(* IEC 61131-3 sources: dvigatel_dorosh/codesys, 10 files *)

(* ---- 00_DUT_MotorTypes.st ---- *)
TYPE E_MotorState :
(
    MOTOR_DISABLED,
    MOTOR_IDLE,
    MOTOR_RAMP,
    MOTOR_WAIT_STOP,
    MOTOR_RUN,
    MOTOR_FAULT
);
END_TYPE

TYPE ST_MotorCommand :
STRUCT
    SpeedRPM : REAL;
    RampSec : REAL;
    Direction : INT; // +1 / -1
    Sequence : WORD;
END_STRUCT
END_TYPE

(* ---- 01_GVL_PC.st ---- *)
VAR_GLOBAL
    // Explicitly map these words into Modbus TCP holding registers in Device Tree.
    // 0..5: PC request. 100..116: PLC telemetry.
    Holding : ARRAY[0..127] OF WORD;

    // Must be commissioned ON SITE; no automatic activation from Ethernet.
    CommissionEnable : BOOL := FALSE;
    ConfigValid : BOOL := FALSE;
    PGFeedbackProven : BOOL := FALSE;
    HardwareSafetyOK : BOOL := FALSE;

    // Assign IO in device mappings, not hard-coded addresses.
    Pt100TemperatureC : REAL;
    Pt100InputValid : BOOL;
END_VAR

(* ---- 07_GVL_DriveIO.st ---- *)
VAR_GLOBAL
    // Link via CODESYS Modbus Serial Device I/O Mapping.
    // NEVER assume default values mean communication is healthy.
    SpeedRaw : WORD;
    StatusRaw : WORD;
    FrequencyRaw : WORD;
    CurrentRaw : WORD;
    FaultCodeRaw : WORD;
    SpeedResponsePulse : BOOL;
    StatusResponsePulse : BOOL;
    DriveReadFresh : BOOL;
    DriveFault : BOOL;

    // Final outputs are NOT directly mapped to a write device in this version.
    // Implement an acknowledged, single-in-flight Modbus RTU scheduler.
    PendingFrequencyWord : WORD;
    PendingControlWord : WORD;
END_VAR

(* ---- 02_FB_Pt100Protection.st ---- *)
FUNCTION_BLOCK FB_Pt100Protection
VAR_INPUT
    TemperatureC : REAL;
    ChannelHealthy : BOOL;
    WarningC : REAL;
    TripC : REAL;
    ResetBelowC : REAL;
    Ack : BOOL;
    LimitsConfigured : BOOL;
END_VAR
VAR_OUTPUT
    Warning : BOOL;
    TripLatched : BOOL;
    Valid : BOOL;
    Permit : BOOL;
END_VAR

Valid := ChannelHealthy AND LimitsConfigured
         AND (ResetBelowC < WarningC)
         AND (WarningC < TripC);
Warning := Valid AND (TemperatureC >= WarningC);

IF (NOT Valid) OR (TemperatureC >= TripC) THEN
    TripLatched := TRUE;
END_IF;

// Acknowledgement alone cannot clear fault if input is missing.
IF Ack AND Valid AND (TemperatureC <= ResetBelowC) THEN
    TripLatched := FALSE;
END_IF;
Permit := Valid AND NOT TripLatched;
END_FUNCTION_BLOCK

(* ---- 03_FB_Heartbeat.st ---- *)
FUNCTION_BLOCK FB_Heartbeat
VAR_INPUT
    Counter : WORD;
    Enable : BOOL;
    CycleSec : REAL;
    TimeoutSec : REAL;
END_VAR
VAR_OUTPUT
    Active : BOOL;
END_VAR
VAR
    Previous : WORD;
    AgeSec : REAL := 10000.0;
    Initialized : BOOL;
END_VAR

IF NOT Enable THEN
    Active := FALSE;
    Initialized := FALSE;
    AgeSec := TimeoutSec;
ELSE
    IF NOT Initialized THEN
        Previous := Counter;
        Initialized := TRUE;
        AgeSec := TimeoutSec;
    ELSIF Counter <> Previous THEN
        Previous := Counter;
        AgeSec := 0.0;
    ELSE
        AgeSec := MIN(10000.0, AgeSec + CycleSec);
    END_IF;
    Active := AgeSec < TimeoutSec;
END_IF;
END_FUNCTION_BLOCK

(* ---- 04_FB_ConfirmedStop.st ---- *)
FUNCTION_BLOCK FB_ConfirmedStop
VAR_INPUT
    EncoderFeedbackProven : BOOL;
    SpeedFresh : BOOL;
    StatusFresh : BOOL;
    DriveReportsStopped : BOOL;
    MeasuredRPM : REAL;
    CycleSec : REAL;
    ThresholdRPM : REAL;
    StableSec : REAL;
END_VAR
VAR_OUTPUT
    Confirmed : BOOL;
END_VAR
VAR
    StableForSec : REAL;
END_VAR

IF EncoderFeedbackProven AND SpeedFresh AND StatusFresh
   AND DriveReportsStopped
   AND (ABS(MeasuredRPM) <= ThresholdRPM)
   AND (StableSec > 0.0) THEN
    StableForSec := MIN(StableSec, StableForSec + CycleSec);
ELSE
    StableForSec := 0.0;
END_IF;
Confirmed := StableForSec >= StableSec AND StableSec > 0.0;
END_FUNCTION_BLOCK

(* ---- 05_FB_MotorMotion.st ---- *)
FUNCTION_BLOCK FB_MotorMotion
VAR_INPUT
    Enable : BOOL;
    InterlocksOK : BOOL;
    CommandPulse : BOOL;
    Command : ST_MotorCommand;
    FaultAck : BOOL;
    StopConfirmed : BOOL;
    CycleSec : REAL;
    MaxRPM : REAL;
    StopTimeoutSec : REAL;
END_VAR
VAR_OUTPUT
    State : E_MotorState := MOTOR_DISABLED;
    ProfileRPM : REAL;             // signed reference
    RunRequest : BOOL;
    ReverseRequest : BOOL;
    StopRequest : BOOL := TRUE;
    FaultLatched : BOOL;
    AcceptedSequence : WORD;
END_VAR
VAR
    Goal : REAL;
    StageStart : REAL;
    StageEnd : REAL;
    StageSec : REAL;
    StageAge : REAL;
    StopAge : REAL;
    PendingReverse : BOOL;
    HeldDirection : INT := 1;
    NewGoal : BOOL;
    ValidCmd : BOOL;
END_VAR

// Device safety must NOT depend on a functioning serial link.
// This output requests a controlled stop; hardware safety is separate.
IF NOT Enable THEN
    State := MOTOR_DISABLED;
    ProfileRPM := 0.0;
    Goal := 0.0;
    PendingReverse := FALSE;
ELSIF NOT InterlocksOK THEN
    FaultLatched := TRUE;
    State := MOTOR_FAULT;
END_IF;

IF State = MOTOR_FAULT THEN
    // Explicit acknowledgement while truly stopped. Does not re-launch.
    IF FaultAck AND InterlocksOK AND StopConfirmed
       AND (Command.SpeedRPM = 0.0) AND NOT CommandPulse THEN
        FaultLatched := FALSE;
        State := MOTOR_IDLE;
        ProfileRPM := 0.0;
        Goal := 0.0;
    END_IF;
ELSIF State = MOTOR_DISABLED THEN
    // Moving from disabled to idle does not accept any pre-existing command.
    IF Enable AND InterlocksOK AND StopConfirmed THEN
        State := MOTOR_IDLE;
    END_IF;
ELSIF Enable AND InterlocksOK THEN
    ValidCmd := (Command.Direction = 1 OR Command.Direction = -1)
            AND (Command.SpeedRPM >= 0.0)
            AND (Command.SpeedRPM <= MaxRPM)
            AND (Command.RampSec >= 0.1)
            AND (Command.RampSec <= 600.0)
            AND (MaxRPM > 0.0);

    NewGoal := CommandPulse AND ValidCmd;
    IF NewGoal THEN
        AcceptedSequence := Command.Sequence;
        Goal := Command.SpeedRPM * INT_TO_REAL(Command.Direction);
        StageSec := Command.RampSec;

        IF State = MOTOR_WAIT_STOP THEN
            // Never cancel physical-stop gate on a new command.
            PendingReverse := (ABS(Goal) > 0.001);
        ELSE
            StageStart := ProfileRPM;
            StageAge := 0.0;
            IF (ABS(ProfileRPM) > 0.001) AND (ABS(Goal) > 0.001)
               AND ((ProfileRPM > 0.0) <> (Goal > 0.0)) THEN
                StageEnd := 0.0;    // reverse: first stop
                PendingReverse := TRUE;
            ELSIF (ABS(ProfileRPM) < 0.001) AND (NOT StopConfirmed)
                  AND (ABS(Goal) > 0.001) THEN
                State := MOTOR_WAIT_STOP;
                StopAge := 0.0;
                PendingReverse := TRUE;
            ELSE
                StageEnd := Goal;
                PendingReverse := FALSE;
                IF ABS(ProfileRPM) < 0.001 AND ABS(Goal) > 0.001 THEN
                    IF Goal < 0.0 THEN HeldDirection := -1;
                    ELSE HeldDirection := 1; END_IF;
                END_IF;
            END_IF;
            IF State <> MOTOR_WAIT_STOP THEN State := MOTOR_RAMP; END_IF;
        END_IF;
    END_IF;

    CASE State OF
        MOTOR_IDLE:
            ProfileRPM := 0.0;

        MOTOR_RAMP:
            StageAge := MIN(StageSec, StageAge + CycleSec);
            ProfileRPM := StageStart +
                 (StageEnd - StageStart) * (StageAge / StageSec);
            IF StageAge >= StageSec THEN
                ProfileRPM := StageEnd;
                IF ABS(StageEnd) <= 0.001 THEN
                    StopAge := 0.0;
                    State := MOTOR_WAIT_STOP;
                ELSE
                    State := MOTOR_RUN;
                END_IF;
            END_IF;

        MOTOR_WAIT_STOP:
            ProfileRPM := 0.0;
            StopAge := StopAge + CycleSec;
            IF StopConfirmed THEN
                IF ABS(Goal) <= 0.001 THEN
                    PendingReverse := FALSE;
                    State := MOTOR_IDLE;
                ELSE
                    IF Goal < 0.0 THEN HeldDirection := -1;
                    ELSE HeldDirection := 1; END_IF;
                    StageStart := 0.0;
                    StageEnd := Goal;
                    StageAge := 0.0;
                    PendingReverse := FALSE;
                    State := MOTOR_RAMP;
                END_IF;
            ELSIF StopAge >= StopTimeoutSec THEN
                FaultLatched := TRUE;
                State := MOTOR_FAULT;
            END_IF;

        MOTOR_RUN:
            ProfileRPM := Goal;
    END_CASE;
END_IF;

// Enforce a stop request for every blocked or waiting state.
RunRequest := (State = MOTOR_RAMP OR State = MOTOR_RUN)
              AND ABS(ProfileRPM) > 0.001
              AND InterlocksOK AND Enable AND NOT FaultLatched;
ReverseRequest := HeldDirection = -1;
StopRequest := NOT RunRequest;
IF State = MOTOR_FAULT OR State = MOTOR_DISABLED THEN
    ProfileRPM := 0.0;
    RunRequest := FALSE;
    StopRequest := TRUE;
END_IF;
END_FUNCTION_BLOCK

(* ---- 06_FB_DriveCommand.st ---- *)
FUNCTION_BLOCK FB_DriveCommand
VAR_INPUT
    ProfileRPM : REAL;
    RunRequest : BOOL;
    ReverseRequest : BOOL;
    StopRequest : BOOL;
    MotorPolePairs : UINT;
    MaximumHz : REAL;
    ConfigurationValid : BOOL;
END_VAR
VAR_OUTPUT
    FrequencyHz : REAL;
    FrequencyWord : WORD;
    ControlWord : WORD;
    Valid : BOOL;
END_VAR

// Feedforward only: true shaft RPM is read from drive.
// This formula does NOT correct asynchronous slip.
Valid := ConfigurationValid AND (MotorPolePairs > 0)
         AND (MaximumHz > 0.0) AND (MaximumHz <= 300.0);
IF NOT Valid THEN
    FrequencyHz := 0.0;
    FrequencyWord := 0;
    ControlWord := 16#0004; // nominal deceleration-stop candidate; verify at bench
ELSE
    FrequencyHz := LIMIT(0.0,
         ABS(ProfileRPM) * UINT_TO_REAL(MotorPolePairs) / 60.0,
         MaximumHz);
    FrequencyWord := REAL_TO_WORD(FrequencyHz * 100.0);
    IF StopRequest OR NOT RunRequest THEN
        ControlWord := 16#0004;
    ELSIF ReverseRequest THEN
        ControlWord := 16#0003;
    ELSE
        ControlWord := 16#0001;
    END_IF;
END_IF;
END_FUNCTION_BLOCK

(* ---- 09_FB_InnovertRTU.st ---- *)
FUNCTION_BLOCK FB_InnovertRTU
VAR_INPUT
    EnablePort : BOOL;
    ComPortNumber : UDINT; // Must be confirmed on PLC200 hardware; zero disables.
    SlaveId : USINT := 1;
    Baudrate : UDINT := 38400;
    EnableWrites : BOOL;   // FALSE until verified commissioning.
    CommandPermitted : BOOL; // Set only after hardware + PG + Pt100 and TCP watchdog.
    SetFrequency : WORD;    // 0.01 Hz units after checking P00.00.
    SetControl : WORD;      // manual confirms 0x0001 forward, 0x0003 reverse, 0x0004 stop.
    CycleSec : REAL := 0.02;
END_VAR
VAR_OUTPUT
    PortActive : BOOL;
    Busy : BOOL;
    Healthy : BOOL;
    LastError : BOOL;
    ErrorCount : UDINT;
    OkCount : UDINT;
    LastOperation : UINT;
    LastFailedOperation : UINT;
    SpeedRaw : WORD;
    StatusRaw : WORD;
    FrequencyRaw : WORD;
    CurrentRaw : WORD;
    FaultRaw : WORD;
    SpeedFresh : BOOL;
    StatusFresh : BOOL;
    TelemetryFresh : BOOL;
    WriteFrequencyAck : BOOL;
    WriteControlAck : BOOL;
    LastWrittenFrequency : WORD;
    LastWrittenControl : WORD;
END_VAR
VAR
    Com : OCL.COM_Control;
    Request : OCL.MB_SerialRequest;
    State : UINT := 0;
    Step : UINT := 0;
    RequestExecute : BOOL;
    FC : OCL.MB_FC;
    RegisterAddress : UINT;
    Payload : WORD;
    StepAge : REAL;
    SpeedAge : REAL := 10000.0;
    StatusAge : REAL := 10000.0;
    CurrentAge : REAL := 10000.0;
    FaultAge : REAL := 10000.0;
    FrequencyAge : REAL := 10000.0;
    PendingFrequency : WORD;
    PendingControl : WORD;
    HadWriteFrequencyAck : BOOL;
    HadWriteControlAck : BOOL;
    ErrorStreak : UINT;
    WriteEligible : BOOL;
    IsWrite : BOOL;
    ReadyPort : BOOL;
END_VAR

// One FB owns one physical port. Never create a second Modbus COM Port
// on the same RS-485 interface in the CODESYS Device Tree.
SpeedFresh := FALSE;
StatusFresh := FALSE;
TelemetryFresh := FALSE;
WriteFrequencyAck := FALSE;
WriteControlAck := FALSE;
LastError := FALSE;
Busy := (State = 20);
SpeedAge := MIN(10000.0, SpeedAge + CycleSec);
StatusAge := MIN(10000.0, StatusAge + CycleSec);
FrequencyAge := MIN(10000.0, FrequencyAge + CycleSec);
CurrentAge := MIN(10000.0, CurrentAge + CycleSec);
FaultAge := MIN(10000.0, FaultAge + CycleSec);

// Avoid opening unspecified COM ports.
ReadyPort := EnablePort AND (ComPortNumber > 0);
Com(
    xEnable := ReadyPort,
    udiComPort := ComPortNumber,
    udiBaudrate := Baudrate,
    udiByteSize := 8,
    eParity := OCL.COM_PARITY.NONE,
    eStopBit := OCL.COM_STOPBIT.ONE
);
PortActive := Com.xActive AND NOT Com.xError;

// Keep one request FB called EVERY PLC task with a rising-edge Execute.
Request(
    xExecute := RequestExecute,
    tTimeout := T#300MS,
    usiRetry := 0,
    hCom := Com.hCom,
    xIsAsciiMode := FALSE,
    usiSlaveId := SlaveId,
    eFuncCode := FC,
    uiDataAddr := RegisterAddress,
    uiDataCount := 1,
    pData := ADR(Payload),
    szSize := SIZEOF(Payload)
);

IF NOT PortActive THEN
    State := 0;
    Step := 0;
    RequestExecute := FALSE;
    ErrorStreak := 0;
    SpeedAge := 10000.0;
    StatusAge := 10000.0;
    Healthy := FALSE;
ELSE
    CASE State OF
    0: // start from read-only polling every time port activates
        Step := 0;
        State := 10;
    10: // choose next operation; readings are serialized.
        RequestExecute := FALSE;
        Payload := 0;
        FC := OCL.MB_FC.READ_HOLDING_REGISTERS;
        IsWrite := FALSE;
        CASE Step OF
        0: RegisterAddress := 16#8107; // RPM
        1: RegisterAddress := 16#8118; // run status
        2: RegisterAddress := 16#8102; // output frequency
        3: RegisterAddress := 16#810A; // output current
        4: RegisterAddress := 16#812B; // fault code
        5:
            // Writing is NEVER enabled by merely connecting the PLC to a PC.
            WriteEligible := EnableWrites AND CommandPermitted
                           AND Healthy AND (SpeedAge < 0.8)
                           AND (StatusAge < 0.8);
            IF WriteEligible THEN
                PendingFrequency := SetFrequency;
                PendingControl := SetControl;
                Payload := PendingFrequency;
                RegisterAddress := 16#0000;
                FC := OCL.MB_FC.WRITE_SINGLE_REGISTER;
                IsWrite := TRUE;
            ELSE
                Step := 0;
                RegisterAddress := 16#8107;
            END_IF;
        6:
            // Cannot write command without a successfully acked frequency write.
            IF HadWriteFrequencyAck AND EnableWrites AND CommandPermitted THEN
                Payload := PendingControl;
                RegisterAddress := 16#8000;
                FC := OCL.MB_FC.WRITE_SINGLE_REGISTER;
                IsWrite := TRUE;
            ELSE
                Step := 0;
                RegisterAddress := 16#8107;
            END_IF;
        ELSE
            Step := 0;
            RegisterAddress := 16#8107;
        END_CASE;
        LastOperation := Step;
        State := 20;
    20: // Hold execute through busy and until Done or Error
        RequestExecute := TRUE;
        IF Request.xDone THEN
            OkCount := OkCount + 1;
            ErrorStreak := 0;
            IF IsWrite THEN
                IF Step = 5 THEN
                    HadWriteFrequencyAck := TRUE;
                    LastWrittenFrequency := PendingFrequency;
                    WriteFrequencyAck := TRUE;
                ELSIF Step = 6 THEN
                    HadWriteControlAck := TRUE;
                    LastWrittenControl := PendingControl;
                    WriteControlAck := TRUE;
                END_IF;
            ELSE
                CASE Step OF
                0:
                    SpeedRaw := Payload;
                    SpeedAge := 0.0;
                    SpeedFresh := TRUE;
                1:
                    StatusRaw := Payload;
                    StatusAge := 0.0;
                    StatusFresh := TRUE;
                2:
                    FrequencyRaw := Payload;
                    FrequencyAge := 0.0;
                3:
                    CurrentRaw := Payload;
                    CurrentAge := 0.0;
                4:
                    FaultRaw := Payload;
                    FaultAge := 0.0;
                END_CASE;
            END_IF;
            State := 30;
        ELSIF Request.xError THEN
            ErrorCount := ErrorCount + 1;
            LastError := TRUE;
            LastFailedOperation := Step;
            ErrorStreak := ErrorStreak + 1;
            HadWriteFrequencyAck := FALSE;
            HadWriteControlAck := FALSE;
            SpeedAge := 10000.0; // fail closed even if status register still has data
            StatusAge := 10000.0;
            State := 30;
        END_IF;
    30: // create falling edge before next request
        RequestExecute := FALSE;
        State := 40;
    40:
        IF Step >= 6 THEN
            Step := 0;
            HadWriteFrequencyAck := FALSE;
        ELSE
            Step := Step + 1;
        END_IF;
        State := 10;
    END_CASE;
END_IF;

Healthy := PortActive AND (ErrorStreak < 3)
           AND (SpeedAge < 0.8) AND (StatusAge < 0.8);
TelemetryFresh := Healthy AND (FrequencyAge < 2.0)
                  AND (CurrentAge < 2.0) AND (FaultAge < 2.0);
Busy := State = 20;
END_FUNCTION_BLOCK

(* ---- 08_PRG_MotorMain.st ---- *)
PROGRAM PRG_MotorMain
VAR
    // Set PLC_PRG task period to 20 ms and verify actual runtime.
    CycleSec : REAL := 0.02;
    TemperatureWarningC : REAL := 0.0; // configure from motor documentation
    TemperatureTripC : REAL := 0.0;
    TemperatureResetC : REAL := 0.0;
    TemperatureLimitsConfigured : BOOL := FALSE;
    MaximumRPM : REAL := 0.0; // set only after mechanical review
    MaximumHz : REAL := 0.0;
    MotorPolePairs : UINT := 0; // expected 2 for 4 poles, verify
    MaxStopWaitSec : REAL := 30.0;

    // These inputs require proven wiring and runtime diagnostics.
    DriveReportsStopped : BOOL := FALSE;
    DriveStatusDecoded : BOOL := FALSE;
    DriveSpeedScalingProven : BOOL := FALSE;
    DriveSpeedSignedRPM : REAL := 0.0;
    DriveResponseAgeSec : REAL := 10000.0;

    RTU : FB_InnovertRTU;
    RTU_ComPort : UDINT := 0; // Set actual PLC200 COM port from hardware diagnostics
    RTU_WriteEnable : BOOL := FALSE; // Must remain FALSE until commissioning
    Temp : FB_Pt100Protection;
    HB : FB_Heartbeat;
    StopCheck : FB_ConfirmedStop;
    Motion : FB_MotorMotion;
    DriveCmd : FB_DriveCommand;

    Cmd : ST_MotorCommand;
    CmdPulse : BOOL;
    LastRequestID : WORD;
    RequestID : WORD;
    RequestDir : INT;
    ValidRequest : BOOL;
    Interlocks : BOOL;
    RunPermitted : BOOL;
    SpeedFresh : BOOL;
    StatusFresh : BOOL;
    TelemetryState : UINT;
    SignedX10 : DINT;
    SignedX10DW : DWORD;
    Ack : BOOL := FALSE; // safety reset must be engineered separately
END_VAR

// Raw RTU communication: use OwenCommunication library; no Modbus COM Port
// device can occupy the same physical RS-485.
RTU(
    EnablePort:=RTU_ComPort > 0,
    ComPortNumber:=RTU_ComPort,
    SlaveId:=1, Baudrate:=38400,
    EnableWrites:=RTU_WriteEnable,
    CommandPermitted:=RunPermitted,
    SetFrequency:=DriveCmd.FrequencyWord,
    SetControl:=DriveCmd.ControlWord,
    CycleSec:=CycleSec
);
GVL_DriveIO.SpeedRaw := RTU.SpeedRaw;
GVL_DriveIO.StatusRaw := RTU.StatusRaw;
GVL_DriveIO.FrequencyRaw := RTU.FrequencyRaw;
GVL_DriveIO.CurrentRaw := RTU.CurrentRaw;
GVL_DriveIO.FaultCodeRaw := RTU.FaultRaw;
GVL_DriveIO.SpeedResponsePulse := RTU.SpeedFresh;
GVL_DriveIO.StatusResponsePulse := RTU.StatusFresh;
GVL_DriveIO.DriveReadFresh := RTU.Healthy;

// WARNING: The following drive-dependent values must be decoded and proven
// from the real IMD222U21E-ENC diagnostics. Not hardwired to TRUE.
// DriveReportsStopped, DriveStatusDecoded, DriveSpeedScalingProven
// and DriveSpeedSignedRPM are commissioning variables.

// Inputs Holding[0..4] must be protected against concurrent partial writes.
// The application accepts ONLY a changed command ID and validated fields.
// For production replace this elementary transaction handling with a
// verified command buffer / consistency token / single writer.
RequestID := GVL_PC.Holding[4];
RequestDir := 0;
IF GVL_PC.Holding[2] = 1 THEN RequestDir := 1; END_IF;
IF GVL_PC.Holding[2] = 2 THEN RequestDir := -1; END_IF;

Cmd.SpeedRPM := WORD_TO_REAL(GVL_PC.Holding[0]) / 10.0;
Cmd.RampSec := WORD_TO_REAL(GVL_PC.Holding[1]) / 10.0;
Cmd.Direction := RequestDir;
Cmd.Sequence := RequestID;
ValidRequest := RequestDir <> 0
    AND Cmd.SpeedRPM >= 0.0 AND Cmd.SpeedRPM <= MaximumRPM
    AND Cmd.RampSec >= 0.1 AND Cmd.RampSec <= 600.0;

CmdPulse := (RequestID <> LastRequestID) AND ValidRequest;
IF RequestID <> LastRequestID THEN LastRequestID := RequestID; END_IF;

Temp(TemperatureC:=GVL_PC.Pt100TemperatureC,
    ChannelHealthy:=GVL_PC.Pt100InputValid,
    WarningC:=TemperatureWarningC, TripC:=TemperatureTripC,
    ResetBelowC:=TemperatureResetC, Ack:=FALSE,
    LimitsConfigured:=TemperatureLimitsConfigured);
HB(Counter:=GVL_PC.Holding[3], Enable:=GVL_PC.CommissionEnable,
   CycleSec:=CycleSec, TimeoutSec:=2.0);

// Freshness: true pulse must be generated on an actual successful RTU response.
IF GVL_DriveIO.DriveReadFresh THEN
    DriveResponseAgeSec := 0.0;
ELSE
    DriveResponseAgeSec := MIN(10000.0, DriveResponseAgeSec + CycleSec);
END_IF;
SpeedFresh := DriveResponseAgeSec < 0.6 AND DriveSpeedScalingProven
              AND GVL_PC.PGFeedbackProven;
StatusFresh := DriveResponseAgeSec < 0.6 AND DriveStatusDecoded;
StopCheck(EncoderFeedbackProven:=GVL_PC.PGFeedbackProven,
    SpeedFresh:=SpeedFresh, StatusFresh:=StatusFresh,
    DriveReportsStopped:=DriveReportsStopped,
    MeasuredRPM:=DriveSpeedSignedRPM, CycleSec:=CycleSec,
    ThresholdRPM:=5.0, StableSec:=0.4);

RunPermitted := GVL_PC.CommissionEnable AND GVL_PC.ConfigValid
    AND GVL_PC.HardwareSafetyOK AND Temp.Permit AND HB.Active
    AND SpeedFresh AND StatusFresh AND NOT GVL_DriveIO.DriveFault;

Interlocks := RunPermitted;
Motion(Enable:=GVL_PC.CommissionEnable AND GVL_PC.ConfigValid,
    InterlocksOK:=Interlocks,
    CommandPulse:=CmdPulse AND HB.Active, Command:=Cmd,
    FaultAck:=FALSE, StopConfirmed:=StopCheck.Confirmed,
    CycleSec:=CycleSec, MaxRPM:=MaximumRPM,
    StopTimeoutSec:=MaxStopWaitSec);
DriveCmd(ProfileRPM:=Motion.ProfileRPM,
    RunRequest:=Motion.RunRequest,
    ReverseRequest:=Motion.ReverseRequest,
    StopRequest:=Motion.StopRequest,
    MotorPolePairs:=MotorPolePairs, MaximumHz:=MaximumHz,
    ConfigurationValid:=GVL_PC.ConfigValid);

// NOT connected to Modbus write requests by default.
// Once RTU scheduler is implemented, it must send frequency and control
// sequentially, verify each acknowledgement, and latch failures.
GVL_DriveIO.PendingFrequencyWord := DriveCmd.FrequencyWord;
GVL_DriveIO.PendingControlWord := DriveCmd.ControlWord;

CASE Motion.State OF
 MOTOR_DISABLED: TelemetryState := 0;
 MOTOR_IDLE: TelemetryState := 1;
 MOTOR_RAMP: TelemetryState := 2;
 MOTOR_WAIT_STOP: TelemetryState := 3;
 MOTOR_RUN: TelemetryState := 4;
 MOTOR_FAULT: TelemetryState := 90;
END_CASE;

GVL_PC.Holding[100] := Motion.AcceptedSequence;
GVL_PC.Holding[101] := UINT_TO_WORD(TelemetryState);
SignedX10 := REAL_TO_DINT(DriveSpeedSignedRPM * 10.0);
SignedX10DW := DINT_TO_DWORD(SignedX10);
GVL_PC.Holding[102] := DWORD_TO_WORD(SHR(SignedX10DW,16));
GVL_PC.Holding[103] := DWORD_TO_WORD(SignedX10DW AND 16#0000FFFF);
IF GVL_PC.Pt100InputValid THEN
 GVL_PC.Holding[104] := INT_TO_WORD(REAL_TO_INT(GVL_PC.Pt100TemperatureC*10.0));
ELSE
 GVL_PC.Holding[104] := 16#7FFF;
END_IF;
GVL_PC.Holding[105] := GVL_DriveIO.FrequencyRaw;
GVL_PC.Holding[106] := GVL_DriveIO.CurrentRaw;
GVL_PC.Holding[107] := GVL_DriveIO.StatusRaw;
GVL_PC.Holding[108] := GVL_DriveIO.FaultCodeRaw;
GVL_PC.Holding[109] := BOOL_TO_WORD(SpeedFresh AND StatusFresh);
GVL_PC.Holding[110] := BOOL_TO_WORD(GVL_PC.PGFeedbackProven);
GVL_PC.Holding[111] := BOOL_TO_WORD(Temp.Permit);
GVL_PC.Holding[112] := BOOL_TO_WORD(StopCheck.Confirmed);
GVL_PC.Holding[113] := DriveCmd.FrequencyWord;
GVL_PC.Holding[114] := DriveCmd.ControlWord;
GVL_PC.Holding[115] := GVL_DriveIO.SpeedRaw;
GVL_PC.Holding[116] := BOOL_TO_WORD(RunPermitted);
END_PROGRAM
